(* IEC 61131-3 sources: sis-interlock-demo/src/POUs/Sis/F_CemCrc, 2 files *)

(* ---- F_CemCrc.decl.st ---- *)
// Назначение: CRC-16/CCITT-FALSE матрицы по 36 байтам: младший и старший байты uiCauseCount,
//             uiEffectCount, затем масок wCauseMask всех 16 следствий (раздел 6.8). Заметить
//             ручную правку сгенерированной конфигурации без генератора (решение D-10).
// Автор:      kr0nsch
// Версия:     0.1.0
// Документ:   docs/DESIGN.md, раздел «6.8 Конфигурация и CRC»
// ВНИМАНИЕ:   код демонстрационный и не предназначен для систем безопасности. Реальная ПАЗ
//             требует определения SIL, сертифицированных аппаратных и программных средств
//             и валидации по ГОСТ Р МЭК 61511.
FUNCTION F_CemCrc : WORD
VAR_IN_OUT CONSTANT
    stCfg : ST_CemCfg;   // конфигурация матрицы
END_VAR
VAR
    wCrc : WORD;         // регистр CRC
    wVal : WORD;         // очередное слово
    uiJ  : UINT;         // индекс следствия
    stEffect : ST_EffectCfg;   // копия столбца
END_VAR

(* ---- F_CemCrc.impl.st ---- *)
wCrc := GVL_Const.CRC16_INIT;

// Слова — младшим байтом вперёд
wVal := UINT_TO_WORD(stCfg.uiCauseCount);
wCrc := F_SisCrc16Byte(wCrc := wCrc, bData := WORD_TO_BYTE(wVal AND GVL_Const.WORD_LOW_BYTE));
wCrc := F_SisCrc16Byte(wCrc := wCrc, bData := WORD_TO_BYTE(SHR(wVal, GVL_Const.BITS_PER_BYTE)));
wVal := UINT_TO_WORD(stCfg.uiEffectCount);
wCrc := F_SisCrc16Byte(wCrc := wCrc, bData := WORD_TO_BYTE(wVal AND GVL_Const.WORD_LOW_BYTE));
wCrc := F_SisCrc16Byte(wCrc := wCrc, bData := WORD_TO_BYTE(SHR(wVal, GVL_Const.BITS_PER_BYTE)));

FOR uiJ := 1 TO GVL_Const.SIS_EFFECTS_MAX DO
    stEffect := stCfg.astEffect[uiJ];
    wVal := stEffect.wCauseMask;
    wCrc := F_SisCrc16Byte(wCrc := wCrc, bData := WORD_TO_BYTE(wVal AND GVL_Const.WORD_LOW_BYTE));
    wCrc := F_SisCrc16Byte(wCrc := wCrc, bData := WORD_TO_BYTE(SHR(wVal, GVL_Const.BITS_PER_BYTE)));
END_FOR

F_CemCrc := wCrc;
